TYPE ST_CylIO :
STRUCT
    xValveWork : BOOL;   // valve AS  (Arbeitsstellung = working position)
    xValveHome : BOOL;   // valve GS  (Grundstellung   = home position)
    xSensWork  : BOOL;   // sensor AS
    xSensHome  : BOOL;   // sensor GS
END_STRUCT
END_TYPE

(* stored: Version 1.1.0.1
   DUT ST_CylIO: Id {518d90e4-fb86-409d-a0a7-1ab318ec328b} *)
